FUNCTION_BLOCK StartFeedPositionHMI (* Basic Function Block Type *)
  (* Standard: 61499-2 *)
  (* Version 0.0, 7/5/2026, Schneider Electric, Template *)
  PACKAGE SE.Nereda;
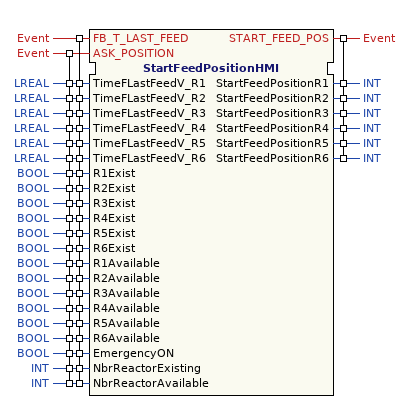
  EVENT_INPUT
    FB_T_LAST_FEED WITH TimeFLastFeedV_R1, TimeFLastFeedV_R2, TimeFLastFeedV_R3, TimeFLastFeedV_R4, TimeFLastFeedV_R5, TimeFLastFeedV_R6, R1Exist, R2Exist, R3Exist, R4Exist, R5Exist, R6Exist, R1Available, R2Available, R3Available, R4Available, R5Available, R6Available, EmergencyON, NbrReactorExisting, NbrReactorAvailable;
    ASK_POSITION WITH TimeFLastFeedV_R1, TimeFLastFeedV_R2, TimeFLastFeedV_R3, TimeFLastFeedV_R4, TimeFLastFeedV_R5, TimeFLastFeedV_R6, R1Exist, R2Exist, R3Exist, R4Exist, R5Exist, R6Exist, R1Available, R2Available, R3Available, R4Available, R5Available, R6Available, EmergencyON, NbrReactorExisting, NbrReactorAvailable;
  END_EVENT
  EVENT_OUTPUT
    START_FEED_POS WITH StartFeedPositionR1, StartFeedPositionR2, StartFeedPositionR3, StartFeedPositionR4, StartFeedPositionR5, StartFeedPositionR6;
  END_EVENT
  VAR_INPUT
    TimeFLastFeedV_R1 : LREAL;
    TimeFLastFeedV_R2 : LREAL;
    TimeFLastFeedV_R3 : LREAL;
    TimeFLastFeedV_R4 : LREAL;
    TimeFLastFeedV_R5 : LREAL;
    TimeFLastFeedV_R6 : LREAL;
    R1Exist : BOOL;
    R2Exist : BOOL;
    R3Exist : BOOL;
    R4Exist : BOOL;
    R5Exist : BOOL;
    R6Exist : BOOL;
    R1Available : BOOL;
    R2Available : BOOL;
    R3Available : BOOL;
    R4Available : BOOL;
    R5Available : BOOL;
    R6Available : BOOL;
    EmergencyON : BOOL;
    NbrReactorExisting : INT;
    NbrReactorAvailable : INT;
  END_VAR
  VAR_OUTPUT
    StartFeedPositionR1 : INT;
    StartFeedPositionR2 : INT;
    StartFeedPositionR3 : INT;
    StartFeedPositionR4 : INT;
    StartFeedPositionR5 : INT;
    StartFeedPositionR6 : INT;
  END_VAR
  VAR
    i : INT := 0;
    ReactorOrder : ARRAY [0..5] OF INT;
    MemoOrder : INT;
    ExAvR1 : BOOL;
    ExAvR2 : BOOL;
  END_VAR
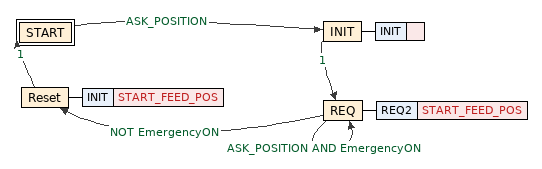
  EC_STATES
    START; (* Initial State *)
    REQ : REQ2 -> START_FEED_POS; (* Normal execution *)
    INIT : INIT;
    Reset : INIT -> START_FEED_POS;
  END_STATES
  EC_TRANSITIONS
    START TO INIT := ASK_POSITION;
    INIT TO REQ := 1;
    Reset TO START := 1;
    REQ TO Reset := NOT EmergencyON;
    REQ TO REQ := ASK_POSITION AND EmergencyON;
  END_TRANSITIONS
  ALGORITHM INIT IN ST:
StartFeedPositionR1 := 0;
StartFeedPositionR2 := 0;
StartFeedPositionR3 := 0;
StartFeedPositionR4 := 0;
StartFeedPositionR5 := 0;
StartFeedPositionR6 := 0;
  END_ALGORITHM
  ALGORITHM REQ2 IN ST:
// Reset all positions at each execution
StartFeedPositionR1 := 0;
StartFeedPositionR2 := 0;
StartFeedPositionR3 := 0;
StartFeedPositionR4 := 0;
StartFeedPositionR5 := 0;
StartFeedPositionR6 := 0;


// ==================================================
// Reactor 1 position
// ==================================================
IF R1Exist AND R1Available THEN

    StartFeedPositionR1 := 1;

    IF R2Exist AND R2Available AND (TimeFLastFeedV_R2 > TimeFLastFeedV_R1) THEN
        StartFeedPositionR1 := StartFeedPositionR1 + 1;
    END_IF;

    IF R3Exist AND R3Available AND (TimeFLastFeedV_R3 > TimeFLastFeedV_R1) THEN
        StartFeedPositionR1 := StartFeedPositionR1 + 1;
    END_IF;

    IF R4Exist AND R4Available AND (TimeFLastFeedV_R4 > TimeFLastFeedV_R1) THEN
        StartFeedPositionR1 := StartFeedPositionR1 + 1;
    END_IF;

    IF R5Exist AND R5Available AND (TimeFLastFeedV_R5 > TimeFLastFeedV_R1) THEN
        StartFeedPositionR1 := StartFeedPositionR1 + 1;
    END_IF;

    IF R6Exist AND R6Available AND (TimeFLastFeedV_R6 > TimeFLastFeedV_R1) THEN
        StartFeedPositionR1 := StartFeedPositionR1 + 1;
    END_IF;

ELSIF R1Exist AND NOT R1Available THEN

    StartFeedPositionR1 := NbrReactorExisting;

END_IF;


// ==================================================
// Reactor 2 position
// ==================================================
IF R2Exist AND R2Available THEN

    StartFeedPositionR2 := 1;

    IF R1Exist AND R1Available AND (TimeFLastFeedV_R1 >= TimeFLastFeedV_R2) THEN
        StartFeedPositionR2 := StartFeedPositionR2 + 1;
    END_IF;

    IF R3Exist AND R3Available AND (TimeFLastFeedV_R3 > TimeFLastFeedV_R2) THEN
        StartFeedPositionR2 := StartFeedPositionR2 + 1;
    END_IF;

    IF R4Exist AND R4Available AND (TimeFLastFeedV_R4 > TimeFLastFeedV_R2) THEN
        StartFeedPositionR2 := StartFeedPositionR2 + 1;
    END_IF;

    IF R5Exist AND R5Available AND (TimeFLastFeedV_R5 > TimeFLastFeedV_R2) THEN
        StartFeedPositionR2 := StartFeedPositionR2 + 1;
    END_IF;

    IF R6Exist AND R6Available AND (TimeFLastFeedV_R6 > TimeFLastFeedV_R2) THEN
        StartFeedPositionR2 := StartFeedPositionR2 + 1;
    END_IF;

ELSIF R2Exist AND NOT R2Available THEN

    StartFeedPositionR2 := NbrReactorExisting;

END_IF;


// ==================================================
// Reactor 3 position
// ==================================================
IF R3Exist AND R3Available THEN

    StartFeedPositionR3 := 1;

    IF R1Exist AND R1Available AND (TimeFLastFeedV_R1 >= TimeFLastFeedV_R3) THEN
        StartFeedPositionR3 := StartFeedPositionR3 + 1;
    END_IF;

    IF R2Exist AND R2Available AND (TimeFLastFeedV_R2 >= TimeFLastFeedV_R3) THEN
        StartFeedPositionR3 := StartFeedPositionR3 + 1;
    END_IF;

    IF R4Exist AND R4Available AND (TimeFLastFeedV_R4 > TimeFLastFeedV_R3) THEN
        StartFeedPositionR3 := StartFeedPositionR3 + 1;
    END_IF;

    IF R5Exist AND R5Available AND (TimeFLastFeedV_R5 > TimeFLastFeedV_R3) THEN
        StartFeedPositionR3 := StartFeedPositionR3 + 1;
    END_IF;

    IF R6Exist AND R6Available AND (TimeFLastFeedV_R6 > TimeFLastFeedV_R3) THEN
        StartFeedPositionR3 := StartFeedPositionR3 + 1;
    END_IF;

ELSIF R3Exist AND NOT R3Available THEN

    StartFeedPositionR3 := NbrReactorExisting;

END_IF;


// ==================================================
// Reactor 4 position
// ==================================================
IF R4Exist AND R4Available THEN

    StartFeedPositionR4 := 1;

    IF R1Exist AND R1Available AND (TimeFLastFeedV_R1 >= TimeFLastFeedV_R4) THEN
        StartFeedPositionR4 := StartFeedPositionR4 + 1;
    END_IF;

    IF R2Exist AND R2Available AND (TimeFLastFeedV_R2 >= TimeFLastFeedV_R4) THEN
        StartFeedPositionR4 := StartFeedPositionR4 + 1;
    END_IF;

    IF R3Exist AND R3Available AND (TimeFLastFeedV_R3 >= TimeFLastFeedV_R4) THEN
        StartFeedPositionR4 := StartFeedPositionR4 + 1;
    END_IF;

    IF R5Exist AND R5Available AND (TimeFLastFeedV_R5 > TimeFLastFeedV_R4) THEN
        StartFeedPositionR4 := StartFeedPositionR4 + 1;
    END_IF;

    IF R6Exist AND R6Available AND (TimeFLastFeedV_R6 > TimeFLastFeedV_R4) THEN
        StartFeedPositionR4 := StartFeedPositionR4 + 1;
    END_IF;

ELSIF R4Exist AND NOT R4Available THEN

    StartFeedPositionR4 := NbrReactorExisting;

END_IF;


// ==================================================
// Reactor 5 position
// ==================================================
IF R5Exist AND R5Available THEN

    StartFeedPositionR5 := 1;

    IF R1Exist AND R1Available AND (TimeFLastFeedV_R1 >= TimeFLastFeedV_R5) THEN
        StartFeedPositionR5 := StartFeedPositionR5 + 1;
    END_IF;

    IF R2Exist AND R2Available AND (TimeFLastFeedV_R2 >= TimeFLastFeedV_R5) THEN
        StartFeedPositionR5 := StartFeedPositionR5 + 1;
    END_IF;

    IF R3Exist AND R3Available AND (TimeFLastFeedV_R3 >= TimeFLastFeedV_R5) THEN
        StartFeedPositionR5 := StartFeedPositionR5 + 1;
    END_IF;

    IF R4Exist AND R4Available AND (TimeFLastFeedV_R4 >= TimeFLastFeedV_R5) THEN
        StartFeedPositionR5 := StartFeedPositionR5 + 1;
    END_IF;

    IF R6Exist AND R6Available AND (TimeFLastFeedV_R6 > TimeFLastFeedV_R5) THEN
        StartFeedPositionR5 := StartFeedPositionR5 + 1;
    END_IF;

ELSIF R5Exist AND NOT R5Available THEN

    StartFeedPositionR5 := NbrReactorExisting;

END_IF;


// ==================================================
// Reactor 6 position
// ==================================================
IF R6Exist AND R6Available THEN

    StartFeedPositionR6 := 1;

    IF R1Exist AND R1Available AND (TimeFLastFeedV_R1 >= TimeFLastFeedV_R6) THEN
        StartFeedPositionR6 := StartFeedPositionR6 + 1;
    END_IF;

    IF R2Exist AND R2Available AND (TimeFLastFeedV_R2 >= TimeFLastFeedV_R6) THEN
        StartFeedPositionR6 := StartFeedPositionR6 + 1;
    END_IF;

    IF R3Exist AND R3Available AND (TimeFLastFeedV_R3 >= TimeFLastFeedV_R6) THEN
        StartFeedPositionR6 := StartFeedPositionR6 + 1;
    END_IF;

    IF R4Exist AND R4Available AND (TimeFLastFeedV_R4 >= TimeFLastFeedV_R6) THEN
        StartFeedPositionR6 := StartFeedPositionR6 + 1;
    END_IF;

    IF R5Exist AND R5Available AND (TimeFLastFeedV_R5 >= TimeFLastFeedV_R6) THEN
        StartFeedPositionR6 := StartFeedPositionR6 + 1;
    END_IF;

ELSIF R6Exist AND NOT R6Available THEN

    StartFeedPositionR6 := NbrReactorExisting;

END_IF;

ASK_POSITION := FALSE;

ReactorOrder[0] := StartFeedPositionR1;
ReactorOrder[1] := StartFeedPositionR2;
ReactorOrder[2] := StartFeedPositionR3;
ReactorOrder[3] := StartFeedPositionR4;
ReactorOrder[4] := StartFeedPositionR5;
ReactorOrder[5] := StartFeedPositionR6;
  END_ALGORITHM
END_FUNCTION_BLOCK
